(*
SPDX-FileCopyrightText: © 2026 Oleksandr Tiutyk <trofimich@gmail.com>
SPDX-License-Identifier: MIT
License: https://opensource.org/license/mit
*)

(*!
<summary>Orders BOOL values described by generic descriptors.</summary>
<description>
Non-null addresses must reference live BOOL storage. TypeClass and Size are not validated and no numeric
conversion is performed. Two null addresses compare equal; one null address sorts before a non-null address.
Descriptors are passed by value; payload remains borrowed and is not modified, cloned, released or retained.
IsMemoryOwner does not affect comparison.
</description>
*)

FUNCTION_BLOCK BoolComparer EXTENDS TOF_Core.Object IMPLEMENTS TOF_Core.IComparer
VAR_STAT
	//! <summary>Class name shared by all instances of this function block.</summary>
	{attribute 'hide'} 
	_ClassName : STRING := __POUNAME();
END_VAR

{attribute 'monitoring' := 'call'}
PROPERTY ClassName : REFERENCE TO STRING
GET
ClassName REF= _ClassName;
END_GET
END_PROPERTY

(*!
<summary>Compares the first operand with the second using this ordering strategy.</summary>
<description>
Non-null addresses must reference live BOOL storage. TypeClass and Size are not validated and no numeric
conversion is performed. Two null addresses compare equal; one null address sorts before a non-null address.
Descriptors are passed by value; payload remains borrowed and is not modified, cloned, released or retained.
IsMemoryOwner does not affect comparison. Descendants cannot replace this standard ordering; implement
IComparer separately for a different ordering strategy.
</description>
*)
//!<param name="first">First descriptor; referenced storage is borrowed for the call.</param>
//!<param name="second">Second descriptor; referenced storage is borrowed for the call.</param>
{attribute "object_name" := "Compare"}
METHOD FINAL Compare : TOF_Core.COMPARISON_RESULT
VAR_INPUT
	first : TOF_Core.GENERIC_VALUE;
	second : TOF_Core.GENERIC_VALUE;
END_VAR
VAR
	leftPointer : POINTER TO BOOL; 
	rightPointer : POINTER TO BOOL; 
END_VAR
IF first.Address = 0 AND_THEN second.Address = 0 THEN
	Compare := TOF_Core.COMPARISON_RESULT.FIRST_EQUAL_TO_SECOND;
	RETURN;
END_IF

IF first.Address = 0 THEN
	Compare := TOF_Core.COMPARISON_RESULT.FIRST_LESS_THAN_SECOND;
	RETURN;	
END_IF

IF second.Address = 0 THEN
	Compare := TOF_Core.COMPARISON_RESULT.FIRST_GREATER_THAN_SECOND;
	RETURN;	
END_IF

leftPointer := first.Address;
rightPointer := second.Address;

IF leftPointer^ < rightPointer^ THEN
	Compare := TOF_Core.COMPARISON_RESULT.FIRST_LESS_THAN_SECOND;
ELSIF leftPointer^ > rightPointer^ THEN
	Compare := TOF_Core.COMPARISON_RESULT.FIRST_GREATER_THAN_SECOND;
ELSE
	Compare := TOF_Core.COMPARISON_RESULT.FIRST_EQUAL_TO_SECOND;	
END_IF
END_METHOD

{attribute 'monitoring' := 'call'}
PROPERTY NamespaceName : REFERENCE TO STRING
GET
NamespaceName REF= CurrentNamespace.Name;
END_GET
END_PROPERTY

{attribute 'monitoring' := 'call'}
PROPERTY SelfSize : ULINT
GET
SelfSize := XSIZEOF(THIS^);
END_GET
END_PROPERTY

END_FUNCTION_BLOCK

(* stored: Version 1.1.0.1
   POU BoolComparer: Id {b24450aa-877e-4dbf-a945-e3d6ba0462d4}, SpecialFunc None
   Property ClassName: Id {4afee12e-0b26-45c8-895f-f54e650a295b}
   Get Get: Id {07ad798a-3c3b-4d44-ba7d-904602efbc06}
   Method Compare: Id {f48eae1f-deb9-4246-bde6-c91900fab6c2}
   Property NamespaceName: Id {57acac9d-d98b-475c-bffd-d8c1f5ad7bb5}
   Get Get: Id {3411fc85-e906-4467-aaf1-f8e6e30593ed}
   Property SelfSize: Id {910da1bd-51d1-4244-858c-df2c2bca4d47}
   Get Get: Id {ece1a941-c310-49ff-ba83-199c5d1387c1} *)
